(* IEC 61131-3 sources: CS_4_Aufzugsteuerung/src/Stations/CP112/Steuerung/Class/_DriveAxisBase (part 2) *)

      16#1B: //27-> PWM setvalue for G-MODE=7 + controlword
        //PWM from -1000 to 1000 for -100% to 100% is preset via SetSpeed
        SyncPara.SetSpeed.size := 2;
        SyncPara.SetSpeed.ptr := #SetValuePtr^.a_SyncValues[x];
        SyncPara.SetSpeed.userinfo := 1;

        SyncPara.ControlWord.size := 2;
        SyncPara.ControlWord.ptr := #SetValuePtr^.a_SyncValues[x] + sizeof(UINT);
        SyncPara.ControlWord.userinfo := 0;

        SyncPara.SetTorque.size := 2;
        SyncPara.SetTorque.ptr := #SetValuePtr^.a_SyncValues[x] + sizeof(UINT);
        SyncPara.SetTorque.userinfo := 0;

    end_case;

  end_for;

END_FUNCTION

FUNCTION VIRTUAL GLOBAL _DriveAxisBase::SetPos::Write
	VAR_INPUT
		input (EAX) 	: DINT;
	END_VAR
	VAR_OUTPUT
		result (EAX) 	: DINT;
	END_VAR

  if (SyncPara.SetPos.ptr <> NIL) & bOnlineFinished then
    SetPos:=input;
    SyncPara.SetPos.ptr^:=input;
  end_if;

 	result := SetPos;

END_FUNCTION

FUNCTION VIRTUAL GLOBAL _DriveAxisBase::SetSpeed::Write
	VAR_INPUT
		input (EAX) 	: DINT;
	END_VAR
	VAR_OUTPUT
		result (EAX) 	: DINT;
	END_VAR

	if bOnlineFinished then
    SetSpeed := Write_SetSpeed(input);  //write value to PDO data, and set possible statusflags.
        end_if;
 	result := SetSpeed;

END_FUNCTION

FUNCTION VIRTUAL GLOBAL _DriveAxisBase::SetCurrent::Write
	VAR_INPUT
		input (EAX) 	: DINT;
	END_VAR
	VAR_OUTPUT
		result (EAX) 	: DINT;
	END_VAR

  if (SyncPara.SetCurrent.ptr <> NIL) & bOnlineFinished then
    SetCurrent:=input;
    if (SyncPara.SetCurrent.size=4) then
      SyncPara.SetCurrent.ptr^:=input;
    elsif (SyncPara.SetCurrent.size=2) then
      if SyncPara.SetCurrent.userinfo = 1 then
        SyncPara.SetCurrent.ptr^$INT:=to_int(input / 10); //because we always get mA and in one case we must send cA
      else
        SyncPara.SetCurrent.ptr^$INT:=to_int(input); //32-Bit-Steuerwort
      end_if;
    end_if;
  end_if;

  result := SetCurrent;

END_FUNCTION

FUNCTION VIRTUAL GLOBAL _DriveAxisBase::ControlWord::Write
	VAR_INPUT
		input (EAX) 	: DS402_Control;
	END_VAR
	VAR_OUTPUT
		result (EAX) 	: DS402_Control;
	END_VAR
  VAR
  	cBuffer : BDINT; //ControlWord Buffer
  END_VAR

  cBuffer := 0; // local variable

  if (SyncPara.ControlWord.ptr <> NIL) & bOnlineFinished then

    if (SyncPara.ControlWord.userinfo=0) then //normal controlword

      cBuffer.1  :=input.EnableOperation;   //DRIVE ENABLE
      cBuffer.2  :=input.ResetFault;        //FAULT RESET
      cBuffer.3  :=input.ManufactureSpec1;  //AMODE2
      cBuffer.4  :=input.ManufactureSpec2;  //KFBRW3
      cBuffer.5  :=input.ManufactureSpec4;  //Output1
      cBuffer.6  :=input.ManufactureSpec5;  //Output2
      cBuffer.7  :=input.ManufactureSpec3;  //KBRAKE
      cBuffer.8  :=input.Reserved1;         //ECHO
      cBuffer.9  :=input.OperationModeSpec1;//SINGLE CAPTURE

      cBuffer:=TorqueCalculation(cBuffer, AxTorqueControl); //cBuffer -> we must add TorqueControl

      SyncPara.ControlWord.ptr^$INT:=to_int(cBuffer);

    elsif(SyncPara.ControlWord.userinfo=1)then

      cBuffer.1 :=input.SwitchOn;
      cBuffer.2 :=input.EnableVoltage;
      cBuffer.3 :=input.QuickStop;
      cBuffer.4 :=input.EnableOperation;    //DRIVE ENABLE
      cBuffer.5 :=input.OperationModeSpec1;
      cBuffer.6 :=input.OperationModeSpec2;
      cBuffer.7 :=input.OperationModeSpec3;
      cBuffer.8 :=input.ResetFault;         //FAULT RESET
      cBuffer.9 :=input.Halt;
      cBuffer.10 :=input.Reserved1;
      cBuffer.11 :=input.Reserved2;
      cBuffer.12 :=input.ManufactureSpec1;  //AMODE2
      cBuffer.13 :=input.ManufactureSpec2;  //KFBRW3
      cBuffer.14 :=input.ManufactureSpec3;  //KBRAKE
      cBuffer.15 :=input.ManufactureSpec4;  //Output1
      cBuffer.16 :=input.ManufactureSpec5;  //Output2

      SyncPara.ControlWord.ptr^$INT:=to_int(cBuffer);

    end_if;

  end_if;

  ControlWord := input;
  result := ControlWord;

END_FUNCTION

FUNCTION VIRTUAL GLOBAL _DriveAxisBase::AxEnable::Write
	VAR_INPUT
		input (EAX) 	: DINT;
	END_VAR
	VAR_OUTPUT
		result (EAX) 	: DINT;
	END_VAR

  if (SyncPara.ControlWord.ptr <> NIL) & bOnlineFinished then
    AxEnable:= Write_Enable( input AND 1 );
  end_if;
  result:=AxEnable;

END_FUNCTION

FUNCTION VIRTUAL GLOBAL _DriveAxisBase::AxErrorQuit::Write
	VAR_INPUT
		input (EAX) 	: DINT;
	END_VAR
	VAR_OUTPUT
		result (EAX) 	: DINT;
	END_VAR

  if SyncPara.ControlWord.ptr & (FirstErrorReset = 0) & bOnlineFinished then

    if (AxError = 1) then

      ErrorQuitHandling(input);

    end_if;

  end_if;

  result := AxErrorQuit;

END_FUNCTION

FUNCTION VIRTUAL GLOBAL _DriveAxisBase::AxTorqueControl::Write
	VAR_INPUT
		input (EAX) 	: UDINT;
	END_VAR
	VAR_OUTPUT
		result (EAX) 	: UDINT;
	END_VAR

  if (SyncPara.SetTorque.ptr <> NIL) & bOnlineFinished then
    SetAxTorque(input);
  end_if;

  result := AxTorqueControl;

END_FUNCTION

FUNCTION _DriveAxisBase::TorqueCalculation
	VAR_INPUT
		cBuffer 	: BDINT;
		input 	  : UDINT;
	END_VAR
	VAR_OUTPUT
		result 	  : BDINT;
	END_VAR
  VAR
  	IReduce   : UDINT;
  END_VAR

  IReduce := ((DRIVEAXIS_TORQUE_LIMITATION_VALUE - input) * 63) / DRIVEAXIS_TORQUE_LIMITATION_VALUE; // calculate the bits for the current reducing

  IReduce := IReduce SHL 10 ;
  cBuffer := cBuffer AND 16#3FF;
  cBuffer+=IReduce$BDINT;

  result:=cBuffer;

END_FUNCTION

//****************************************************************************************************\\
//**################################################################################################**\\
//**************************** everything for getting the actual values!! ****************************\\
//**################################################################################################**\\
//****************************************************************************************************\\

FUNCTION VIRTUAL GLOBAL _DriveAxisBase::GetSynchronPara
  VAR
  	x:SINT;
    SetAVALTT:HSINT;
  END_VAR

  ActValuePtr := DriveMng.GetAxisRdPtr(usAxisIndex); // Zeiger auf die Sollwerte von der Struktur t_ReadValuePtr

  for x:=4 to 0 by -1 do
    SetAVALTT:=ActValues[x];

    case SetAVALTT of

      16#01: //1 -> I-N
        SyncPara.ActSpeed.ptr:=#ActValuePtr^.a_SyncValues[x];
        SyncPara.ActSpeed.size:=4;
        SyncPara.ActSpeed.userinfo:=0;

      16#02: //2 -> I-NFILT
        SyncPara.ActSpeed.ptr:=#ActValuePtr^.a_SyncValues[x];
        SyncPara.ActSpeed.size:=4;
        SyncPara.ActSpeed.userinfo:=0;

//      16#03:
//
//        SyncPara.SetPos

      16#05: //5 -> I-IQ
        SyncPara.ActCurrent.ptr:=#ActValuePtr^.a_SyncValues[x];
        SyncPara.ActCurrent.size:=4;
        SyncPara.ActCurrent.userinfo:=0;

      16#07: //7 -> I-POS
        SyncPara.ActPos.ptr:=#ActValuePtr^.a_SyncValues[x];
        SyncPara.ActPos.size:=4;
        SyncPara.ActPos.userinfo:=0;

      16#09: //9 -> I-PE
        SyncPara.Xw.ptr:=#ActValuePtr^.a_SyncValues[x];
        SyncPara.Xw.size:=4;
        SyncPara.Xw.userinfo:=0;

      16#0A: //10 -> I-IQ + stateword (cA!)
        SyncPara.ActCurrent.ptr:=#ActValuePtr^.a_SyncValues[x];
        SyncPara.ActCurrent.size:=2;
        SyncPara.ActCurrent.userinfo:=1;

        SyncPara.StateWord.ptr:=#ActValuePtr^.a_SyncValues[x]+sizeof(UINT);
        SyncPara.StateWord.size:=2;
        SyncPara.StateWord.userinfo:=0;

      16#0E: //14 -> I-PE + stateword
        SyncPara.Xw.ptr:=#ActValuePtr^.a_SyncValues[x];
        SyncPara.Xw.size:=2;
        SyncPara.Xw.userinfo:=0;

        SyncPara.StateWord.ptr:=#ActValuePtr^.a_SyncValues[x]+sizeof(UINT);
        SyncPara.StateWord.size:=2;
        SyncPara.StateWord.userinfo:=0;

      16#14: //20 -> Current in Promille + stateword
        SyncPara.ActCurrent.ptr:=#ActValuePtr^.a_SyncValues[x];
        SyncPara.ActCurrent.size:=2;
        SyncPara.ActCurrent.userinfo:=0;

        SyncPara.StateWord.ptr:=#ActValuePtr^.a_SyncValues[x]+sizeof(UINT);
        SyncPara.StateWord.size:=2;
        SyncPara.StateWord.userinfo:=1;

      16#15: //21 -> I-POS 2 position of optional encoder
        if (SyncPara.ActPos.ptr = NIL) then
          SyncPara.ActPos.ptr:=#ActValuePtr^.a_SyncValues[x];
          SyncPara.ActPos.size:=4;
          SyncPara.ActPos.userinfo:=0;
        end_if;

      16#17: //23 -> digital inputs + stateword
        SyncPara.DigInputs.ptr:=#ActValuePtr^.a_SyncValues[x];
        SyncPara.DigInputs.size:=8; //no inputs
        SyncPara.DigInputs.userinfo:=0;

        SyncPara.StateWord.ptr:=#ActValuePtr^.a_SyncValues[x]+sizeof(UINT);
        SyncPara.StateWord.size:=2;
        SyncPara.StateWord.userinfo:=0;

      16#1C: //28 -> MultiTurn Pos VSDC151
        SyncPara.ActPos.ptr:=#ActValuePtr^.a_SyncValues[x];
        SyncPara.ActPos.size:=4;
        SyncPara.ActPos.userinfo:=0;

    end_case;

  end_for;

END_FUNCTION

FUNCTION VIRTUAL GLOBAL _DriveAxisBase::ActPos::Read
	VAR_OUTPUT
		output (EAX) 	: DINT;
	END_VAR

  if (SyncPara.ActPos.ptr <> NIL) & bOnlineFinished then
    ActPos:=SyncPara.ActPos.ptr^;
  else
    ActPos:=0;
  end_if;

  output := ActPos;

END_FUNCTION

FUNCTION VIRTUAL GLOBAL _DriveAxisBase::ActSpeed::Read
	VAR_OUTPUT
		output (EAX) 	: DINT;
	END_VAR

  if (SyncPara.ActSpeed.ptr <> NIL) & bOnlineFinished then
    ActSpeed:=SyncPara.ActSpeed.ptr^;
  else
    ActSpeed:=0;
  end_if;

  output := ActSpeed;

END_FUNCTION

FUNCTION VIRTUAL GLOBAL _DriveAxisBase::ActCurrent::Read
	VAR_OUTPUT
		output (EAX) 	: DINT;
	END_VAR

  if (SyncPara.ActCurrent.ptr <> NIL) & bOnlineFinished then
    if SyncPara.ActCurrent.size = 4 then
      ActCurrent:=SyncPara.ActCurrent.ptr^;

    elsif SyncPara.ActCurrent.size = 2 then
      if SyncPara.ActCurrent.userinfo = 1 then
        ActCurrent := to_dint(SyncPara.ActCurrent.ptr^$INT) * 10; //because we want to see mA and not cA
      else
        ActCurrent := to_dint(SyncPara.ActCurrent.ptr^$INT);
      end_if;
    end_if;
  else
    ActCurrent:=0;
  end_if;

  output := ActCurrent;

END_FUNCTION

FUNCTION VIRTUAL GLOBAL _DriveAxisBase::ActXw::Read
	VAR_OUTPUT
		output (EAX) 	: DINT;
	END_VAR

  if (SyncPara.Xw.ptr <> NIL) & bOnlineFinished then
    if SyncPara.Xw.size = 4 then
      ActXw:=SyncPara.Xw.ptr^;
    elsif SyncPara.Xw.size = 2 then
      ActXw := to_dint(SyncPara.Xw.ptr^$INT);
    end_if;
  else
    ActXw:=0;
  end_if;

  output := ActXw;

END_FUNCTION

FUNCTION VIRTUAL GLOBAL _DriveAxisBase::StateWord::Read
	VAR_OUTPUT
		output (EAX) 	: DS402_State;
	END_VAR
  VAR
  	sBuffer : BDINT; //StateWord Buffer
  END_VAR

  if (SyncPara.StateWord.ptr <> NIL) & bOnlineFinished then
    sBuffer := SyncPara.StateWord.ptr^$BDINT; //normales Statuswort

    if (SyncPara.StateWord.userinfo=0) then
      StateWord.ReadyToSwitchOn     :=  sBuffer.1;  //READY TO SWITCH ON
      StateWord.SwitchedOn          :=  sBuffer.2;  //EXT ENABLE LOCKED&ENABLE
      StateWord.OperationEnabled    :=  sBuffer.3;  //OPERATION_ENABLE
      StateWord.Fault               :=  sBuffer.4;  //ERROR
      StateWord.Warning             :=  sBuffer.5;  //WARNING
      StateWord.Remote              :=  sBuffer.6;  //PLL Bit0
      StateWord.VoltageEnabled      :=  sBuffer.7;  //PLL Bit1
      StateWord.SwitchOnDisabled    :=  sBuffer.8;  //ECHO
      StateWord.OperationModeSpec1  :=  sBuffer.9;  //Capture Toggle Bit (I-CAP)
      StateWord.OperationModeSpec2  :=  sBuffer.10; //Capture 4 Toggle Bit (I-CAP4)
      StateWord.InternalLimitActive :=  sBuffer.11; //MULTITURN REVOLUTION ERROR
      StateWord.ManufactureSpec1    :=  sBuffer.12; //Digital Input 1
      StateWord.ManufactureSpec2    :=  sBuffer.13; //Digital Input 2
      StateWord.ManufactureSpec3    :=  sBuffer.14; //Digital Input 3
      StateWord.QuickStop           :=  sBuffer.15; //Digital Input 4
      StateWord.TargetReached       :=  sBuffer.16; //Digital Input 5

    elsif(SyncPara.StateWord.userinfo=1) then
      StateWord.ReadyToSwitchOn     :=  sBuffer.1;  //READY TO SWITCH ON
      StateWord.SwitchedOn          :=  sBuffer.2;  //EXT.ENABLE=LOCKED&ENABLE
      StateWord.OperationEnabled    :=  sBuffer.3;  //OPERATION_ENABLE
      StateWord.Fault               :=  sBuffer.4;  //ERROR
      StateWord.Warning             :=  sBuffer.5;  //WARNING
      StateWord.QuickStop           :=  sBuffer.6;
      StateWord.SwitchOnDisabled    :=  sBuffer.7;
      StateWord.VoltageEnabled      :=  sBuffer.8;
      StateWord.ManufactureSpec1    :=  sBuffer.9;
      StateWord.ManufactureSpec2    :=  sBuffer.10;
      StateWord.TargetReached       :=  sBuffer.11;
      StateWord.ManufactureSpec3    :=  sBuffer.12;
      StateWord.OperationModeSpec1  :=  sBuffer.13;
      StateWord.OperationModeSpec2  :=  sBuffer.14;
      StateWord.Remote              :=  sBuffer.15; //PLL nicht eingerastet
      StateWord.InternalLimitActive :=  sBuffer.16; //MULTITURN REVOLUTION ERROR
    end_if;

  else
    StateWord := 0;
  end_if;

  output := StateWord;

END_FUNCTION

FUNCTION VIRTUAL GLOBAL _DriveAxisBase::AxError::Read
	VAR_OUTPUT
		output (EAX) : DINT;
	END_VAR

  //Error of Axis gets only shown, if Axis is Online
  if bOnlineFinished then
    AxError := GetAxError();
  else
    AxError := 0;
  end_if;

  output := AxError;

END_FUNCTION

FUNCTION _DriveAxisBase::LoadDrivePara
  VAR
    pTabAdress : ^DINT;
    TabLength   : DINT;
  END_VAR

  // load the parameter data to the para objects
  case DriveInitType of

    _SDDSTDTABLE :

     pTabAdress := GetTabAdress(TabType:= 0, bdSettings.bSendMPara, #TabLength);
     SetListToParObj(pData:= (pTabAdress)$^DINT, udLen:=TabLength$UDINT);

    _SDDL2TABLE :
    // load the data of the table
      pTabAdress := GetTabAdress(TabType:= 1, bdSettings.bSendMPara, #TabLength);
      SetListToParObj(pData:= (pTabAdress)$^DINT, udLen:=TabLength$UDINT);

    _SDDRAMEX,
    _SDDFILE :
      pSDDData$^void := DriveAxisSet.GetMemPtr();
      if pSDDData <> NIL then
        // load the data of the memory
        SetListToParObj(pData:= (pSDDData$DINT + pSDDData^.AxOffset)$^DINT, udLen:=pSDDData^.AxLength);
      end_if;

  end_case;

END_FUNCTION

FUNCTION _DriveAxisBase::SetListToParObj
	VAR_INPUT
		pData 	: ^DINT;
		udLen 	: UDINT;
	END_VAR
	VAR_OUTPUT
		retcode 	: BOOL;
	END_VAR
  VAR
    pHlp          : ^DINT;
    x             : UDINT;
    pThisNewInst  : ^void;
    usParaNr      : USINT;
    ParaValue     : DINT;
    UserPara      : CmdStruct;
    UserResult    : Results;
  END_VAR

  retcode := FALSE;

  //hier konnte es zu einem Problem kommen kann wenn pThisNewInst nicht init war.
  pThisNewInst := NIL; //BleErn 19.08.2010 11:27

  if (bdSettings.bAxSetPara = FALSE) | (pData = NIL) then
    return;
  end_if;

  x := 0;
  pHlp := pData;

  while x < udLen do

    usParaNr := pHlp^$USINT;
    pHlp += sizeof(USINT);
    x += sizeof(USINT);

    if usParaNr <= MAX_MOTOR_PARA then
      pThisNewInst$DINT := AxSetPara[IDX_MOTOR_PARA];
    elsif usParaNr <= MAX_DRIVE_PARA then
      pThisNewInst$DINT := AxSetPara[IDX_DRIVE_PARA];
    elsif usParaNr <= MAX_CURRENT_PARA then
      pThisNewInst$DINT := AxSetPara[IDX_CURRENT_PARA];
    elsif usParaNr <= MAX_VEL_PARA then
      pThisNewInst$DINT := AxSetPara[IDX_VEL_PARA];
    elsif usParaNr <= MAX_POS_PARA then
      pThisNewInst$DINT := AxSetPara[IDX_POS_PARA];
    elsif usParaNr <= MAX_FD_PARA then
      pThisNewInst$DINT := AxSetPara[IDX_FD_PARA];
    elsif usParaNr <= MAX_APPLI_PARA then
      pThisNewInst$DINT := AxSetPara[IDX_APPLI_PARA];
    elsif usParaNr <= MAX_ERRORHANDLING then
      pThisNewInst$DINT := AxSetPara[IDX_ERRORHANDLING];
    end_if;

    ParaValue := pHlp^$DINT;
    if pThisNewInst <> NIL then
      UserPara.uiCmd := SDD_REFRESH_SETPARA;
      UserPara.aPara[0] := to_dint(usParaNr);
      UserPara.aPara[1] := ParaValue;
      pThisNewInst$^VirtualBase^.NewInst(#UserPara, #UserResult);
    end_if;

    pHlp += sizeof(UDINT);
    x += sizeof(UDINT);

  end_while;

END_FUNCTION

FUNCTION VIRTUAL GLOBAL _DriveAxisBase::SDDProcess
  VAR
    tmpStr : array [0..20] of char;
    retcode : iprStates;
    dError : DINT;
  END_VAR

  //SA 23391 - ObeChr: Wait for Online before starting SDDCmdInterface
  if Online = 1 then

    case SDDCmdIntfc of

    _SDDIDLE :
      // do nothing

    _SDDREADALL :
      if bdSettings.bStartRead = FALSE then
        bdSettings.bStartRead := TRUE;
        // check if a read is possible
        if ChkParaRead(0) = FALSE then
          SDDCmdIntfc := _SDDIDLE;
        else
          ParaReadProc();
        end_if;
      else
        // überprüfen ob alle Parameter schon vorhanden sind
        ParaReadProc();
        if (bdSettings.bReadAxFin = TRUE) then
          SDDCmdIntfc := _SDDIDLE;
          bdSettings.bStartRead := FALSE;
        end_if;
      end_if;

    _SDDINIT :

      if (AxEnable = 0)  then
        if OldSDDCmdIntfc <> SDDCmdIntfc then
          DriveMng.InitDrive(0); // start the initialisation of the drive
          Init_Again:=true;
          //bdSettings.bDriveInitialized:=true;
        end_if;
      else
        SDDCmdIntfc := _SDDIDLE;
      end_if;

    _SDDURINIT :

      if (AxEnable = 0) then
        if OldSDDCmdIntfc <> SDDCmdIntfc then
          DriveMng.InitDrive(1); // start the initialisation of the drive
          InitASyncPara(); // initialize the structure
          Init_Again:=true;
        end_if;
      else
        SDDCmdIntfc := _SDDIDLE;
      end_if;

    _SDDEXDATA,
    _SDDEXDATAXML:

      // only if a object of the correct class is connected
      if DriveAxisSet.ChkFileHandle() then

        if OldSDDCmdIntfc <> SDDCmdIntfc then
          pSDDData$^void := DriveAxisSet.GetMemPtr();

          // Always Call SetDriveType incause GetDriveTypeStr fails or an older Version of _DriveFileHandling is used
          DriveAxisSet.SetDriveType(eDriveType:=GetDriveType());

          _strcpy(#pSDDData^.AxName[0],#szObjName[0]); //here the name of the object is set to the struct

          // Set tmpStr to 0 incase GetDriveTypeStr does not return a valid string.
          tmpStr[0] := 0;
          DriveMng.GetDriveTypeStr(eDriveType:=GetDriveType(), pDriveTypeStr:=#tmpStr[0], DriveTypeStrSize:=sizeof(tmpStr) );
          if tmpStr[0] then
            DriveAxisSet.SetDriveTypeStr(pDriveTypeStr:= #tmpStr[0]);
          end_if;
          DriveAxisSet.SetUserSSDCmd(SDDCmdIntfc, pSDDData);

        else
          SDDCmdIntfc := DriveAxisSet.GetUserSSDCmd();
        end_if;
      else
        LogError(pMsg:="@06F3 (_DriveAxisBase::SDDProcess) Failed export drive parameters. Check if client 'FileHandle' is connected.");
        SDDCmdIntfc := _SDDERROR;
      end_if;

    _SDDIMDATAXML:

      if DriveAxisSet.ChkFileHandle() then

        if OldSDDCmdIntfc <> SDDCmdIntfc then
          pSDDData$^void := DriveAxisSet.GetMemPtr();

          _strcpy(#pSDDData^.AxName[0],#szObjName[0]); //here the name of the object is set to the struct
          DriveAxisSet.SetUserSSDCmd(SDDCmdIntfc, pSDDData);

        else

          if DriveAxisSet.GetUserSSDCmd() = _SDDIDLE then
            // Read xml file done

            // Insert Crc into the imported Data
            pSDDData^.udCRC32 := DriveAxisSet.CalcCRC32((pSDDData + sizeof(UDINT))$^UDINT, pSDDData^.udLen - sizeof(UDINT));

            // now save all parameters in the SRAM / FILE
            if DriveInitType = _SDDRAMEX then
              pSDDData$^void := DriveAxisSet.GetMemPtr();
              DriveAxisSet.SaveRamExData(pData:= pSDDData, udLen:= pSDDData^.udLen, udOffset:= 0);

            elsif DriveInitType = _SDDFILE then
              pSDDData$^void := DriveAxisSet.GetMemPtr();
              DriveAxisSet.SaveRamFileData(pData:= pSDDData, udLen:= pSDDData^.udLen, udOffset:= 0);

            end_if;

            // Use _SDDINIT to tranfer Parametera from ramfile/sram to drive
            SDDCmdIntfc := _SDDINIT;  // Set after SaveRamExData, SaveRamFileData because Filehandling may suspend task

            return; // Return needed here so that _SDDINIT is registered as a new command
          end_if;

        end_if;
      else
        LogError(pMsg:="@06F5 (_DriveAxisBase::SDDProcess) Failed import drive parameters. Check if client 'FileHandle' is connected.");
        SDDCmdIntfc := _SDDERROR;
      end_if;

      _SDDEXLOGFILE:

        // First call since SDDCmdIntfc was set.
        if OldSDDCmdIntfc <> SDDCmdIntfc then

          retcode := DriveMng.GetLogFile(pDestinationDPNE:=NIL, pdError:=#dError);

          if retcode = ERROR then

            LogValue("@0846 (_DriveAxisBase::SDDProcess) Failed to start read logfile. Error code: -0x{0}", (-dError)$UDINT);
            SDDCmdIntfc := _SDDERROR;

          end_if;

        else

          retcode := DriveMng.GetFileState(pdError:=#dError);

          if retcode = READY then

            SDDCmdIntfc := _SDDIDLE;

          elsif retcode = ERROR then

            LogValue("@0847 (_DriveAxisBase::SDDProcess) Failed read logfile. Error code: -0x{0}", (-dError)$UDINT);
            SDDCmdIntfc := _SDDERROR;

          end_if;

        end_if;

    end_case;

    OldSDDCmdIntfc := SDDCmdIntfc;

  end_if;

END_FUNCTION

FUNCTION VIRTUAL GLOBAL _DriveAxisBase::SDDCmdIntfc::Write
	VAR_INPUT
		input (EAX) 	: _SDDUSERCMD;
	END_VAR
	VAR_OUTPUT
		result (EAX) 	: _SDDUSERCMD;
	END_VAR

  if ((SDDCmdIntfc = _SDDIDLE) |
      (SDDCmdIntfc = _SDDERROR)) then
    SDDCmdIntfc := input;
    result := SDDCmdIntfc;
  else
    result$DINT := ACCESS_DENIED;
  end_if;

END_FUNCTION

FUNCTION _DriveAxisBase::ChkParaRead
	VAR_INPUT
		ChkType 	: DINT;
	END_VAR
	VAR_OUTPUT
		retcode 	: BOOL;
	END_VAR

  retcode := FALSE;

  case ChkType of
  0 : // check if a reading command is allowed

    bdSettings.bReadAx := FALSE;

    bdSettings.bReadAxFin := FALSE;

    if (bdSettings.bAxSetPara = TRUE)then
      bdSettings.bReadAx := TRUE;
      ParaReadCmdAx := 1;
      retcode := TRUE;
    else
      bdSettings.bReadAxFin := TRUE;
    end_if;

  1 : // check if we can send the next reading commands
    if ParaReadCmdAx = 2 then
      if AxASyncPara.ActEntries < 10 then
        retcode := TRUE;
      end_if;
    end_if;

  end_case;

END_FUNCTION

FUNCTION _DriveAxisBase::ParaReadProc
  VAR
    dValue      : DINT;
    pThis       : ^void;
    i           : DINT;
    UserPara    : CmdStruct;
    UserResult  : Results;
  END_VAR
        // Start laden aller Parameter vom Drive
        // folgender Ablauf :
        // 1. Es wird für jede Achse die Anforderung in den Ringbuffer geschrieben (30mal).(Eigene Kennung erforderlich ?);
        // 2. Warten bis nur mehr 10 Einträge vorhanden sind, und dann die nächsten Einträge absetzen
        // 3. wenn alle Einträge abgesetzt sind, (letzter Eintrag muss eine extra Kennung haben), wird überprüft wann alle Daten vorhanden sind
        // 4. Wenn ein Wert eines Parameters ankommt, wird dieser in den Speicher geschrieben, dies ist abhängig von der Sicherungsauswahl. Ist eine Tabelle ausgewählt
        //    werden die Daten sofort an die Parameterklassen gesendet, sind keine Parameterobjekte vorhanden, so wird der Vorgang gar nicht durchgeführt.
        // 5. Wenn der letzte Wert des Parameters kommt, wird die Chksumme neu berechnet, die Daten weggesichert, und die Parameterobjekte aktualisiert

  dValue := 0;

 if bdSettings.bReadAx = TRUE then
    case ParaReadCmdAx of

    0 : //idle step

    1 : // set the first entries in the buffer
      // set the info busy to all para classes
      UserPara.uiCmd := SDD_ASYNC_BUSY;

      for i := IDX_MOTOR_PARA to IDX_ERRORHANDLING do
        pThis$DINT := AxSetPara[i];
        if pThis <> NIL then
          // Set the state BUSY
          pThis$^VirtualBase^.NewInst(#UserPara, #UserResult);
        end_if;
      end_for;

      if AxSetPara[IDX_MOTOR_PARA] <> 0 then
        pThis$DINT := AxSetPara[IDX_MOTOR_PARA];

        AddASyncEntry(usParaNr:= SDD_M_NAME1, usRdWr:= 0, dValue:= dValue, pThisObj:= pThis, usEntry:= 1);
        AddASyncEntry(usParaNr:= SDD_M_NAME2, usRdWr:= 0, dValue:= dValue, pThisObj:= pThis, usEntry:= 1);
        AddASyncEntry(usParaNr:= SDD_M_NAME3, usRdWr:= 0, dValue:= dValue, pThisObj:= pThis, usEntry:= 1);
        AddASyncEntry(usParaNr:= SDD_M_INULL, usRdWr:= 0, dValue:= dValue, pThisObj:= pThis, usEntry:= 1);
        AddASyncEntry(usParaNr:= SDD_M_IPEAK, usRdWr:= 0, dValue:= dValue, pThisObj:= pThis, usEntry:= 1);
        AddASyncEntry(usParaNr:= SDD_M_NMAX, usRdWr:= 0, dValue:= dValue, pThisObj:= pThis, usEntry:= 1);
        AddASyncEntry(usParaNr:= SDD_M_POL, usRdWr:= 0, dValue:= dValue, pThisObj:= pThis, usEntry:= 1);
        AddASyncEntry(usParaNr:= SDD_M_TORQUE, usRdWr:= 0, dValue:= dValue, pThisObj:= pThis, usEntry:= 1);
        AddASyncEntry(usParaNr:= SDD_M_L, usRdWr:= 0, dValue:= dValue, pThisObj:= pThis, usEntry:= 1);
        AddASyncEntry(usParaNr:= SDD_M_R, usRdWr:= 0, dValue:= dValue, pThisObj:= pThis, usEntry:= 1);
        AddASyncEntry(usParaNr:= SDD_M_J, usRdWr:= 0, dValue:= dValue, pThisObj:= pThis, usEntry:= 1);
        AddASyncEntry(usParaNr:= SDD_M_TYPE, usRdWr:= 0, dValue:= dValue, pThisObj:= pThis, usEntry:= 1);
        AddASyncEntry(usParaNr:= SDD_M_RPOL, usRdWr:= 0, dValue:= dValue, pThisObj:= pThis, usEntry:= 1);
        AddASyncEntry(usParaNr:= SDD_M_ROFF, usRdWr:= 0, dValue:= dValue, pThisObj:= pThis, usEntry:= 1);
        AddASyncEntry(usParaNr:= SDD_M_RPULSE, usRdWr:= 0, dValue:= dValue, pThisObj:= pThis, usEntry:= 1);
        AddASyncEntry(usParaNr:= SDD_M_RTEMP, usRdWr:= 0, dValue:= dValue, pThisObj:= pThis, usEntry:= 1);
        AddASyncEntry(usParaNr:= SDD_M_SER, usRdWr:= 0, dValue:= dValue, pThisObj:= pThis, usEntry:= 1);
        AddASyncEntry(usParaNr:= SDD_M_BRAKE, usRdWr:= 0, dValue:= dValue, pThisObj:= pThis, usEntry:= 1);
        AddASyncEntry(usParaNr:= SDD_M_IFWEAK, usRdWr:= 0, dValue:= dValue, pThisObj:= pThis, usEntry:= 1);
        AddASyncEntry(usParaNr:= SDD_M_BRDIS, usRdWr:= 0, dValue:= dValue, pThisObj:= pThis, usEntry:= 1);
        AddASyncEntry(usParaNr:= SDD_M_BREN, usRdWr:= 0, dValue:= dValue, pThisObj:= pThis, usEntry:= 1);
        AddASyncEntry(usParaNr:= SDD_M_IMAG, usRdWr:= 0, dValue:= dValue, pThisObj:= pThis, usEntry:= 1);
        AddASyncEntry(usParaNr:= SDD_M_TROT, usRdWr:= 0, dValue:= dValue, pThisObj:= pThis, usEntry:= 1);
        AddASyncEntry(usParaNr:= SDD_M_UN, usRdWr:= 0, dValue:= dValue, pThisObj:= pThis, usEntry:= 1);
        AddASyncEntry(usParaNr:= SDD_M_UBOOST, usRdWr:= 0, dValue:= dValue, pThisObj:= pThis, usEntry:= 1);
        AddASyncEntry(usParaNr:= SDD_M_KN, usRdWr:= 0, dValue:= dValue, pThisObj:= pThis, usEntry:= 1);
      end_if;

      if AxSetPara[IDX_DRIVE_PARA] <> 0 then
        pThis$DINT := AxSetPara[IDX_DRIVE_PARA];
        AddASyncEntry(usParaNr:= SDD_G_MODE, usRdWr:= 0, dValue:= dValue, pThisObj:= pThis, usEntry:= 1);
        AddASyncEntry(usParaNr:= SDD_G_CETIME, usRdWr:= 0, dValue:= dValue, pThisObj:= pThis, usEntry:= 1);
        AddASyncEntry(usParaNr:= SDD_G_VMAINS, usRdWr:= 0, dValue:= dValue, pThisObj:= pThis, usEntry:= 1);
        AddASyncEntry(usParaNr:= SDD_G_VBUSM, usRdWr:= 0, dValue:= dValue, pThisObj:= pThis, usEntry:= 1);
        AddASyncEntry(usParaNr:= SDD_G_VBUSM, usRdWr:= 0, dValue:= dValue, pThisObj:= pThis, usEntry:= 1);
        AddASyncEntry(usParaNr:= SDD_G_MTEMPK, usRdWr:= 0, dValue:= dValue, pThisObj:= pThis, usEntry:= 1);
        AddASyncEntry(usParaNr:= SDD_G_MTEMPE, usRdWr:= 0, dValue:= dValue, pThisObj:= pThis, usEntry:= 1);
        AddASyncEntry(usParaNr:= SDD_G_PWM, usRdWr:= 0, dValue:= dValue, pThisObj:= pThis, usEntry:= 1);
        AddASyncEntry(usParaNr:= SDD_G_DELAY, usRdWr:= 0, dValue:= dValue, pThisObj:= pThis, usEntry:= 1);
        AddASyncEntry(usParaNr:= SDD_G_FTEMP, usRdWr:= 0, dValue:= dValue, pThisObj:= pThis, usEntry:= 1);
        AddASyncEntry(usParaNr:= SDD_G_EMRAMP, usRdWr:= 0, dValue:= dValue, pThisObj:= pThis, usEntry:= 1);
        AddASyncEntry(usParaNr:= SDD_G_MASKE1, usRdWr:= 0, dValue:= dValue, pThisObj:= pThis, usEntry:= 1);
        AddASyncEntry(usParaNr:= SDD_G_MASKE2, usRdWr:= 0, dValue:= dValue, pThisObj:= pThis, usEntry:= 1);
        AddASyncEntry(usParaNr:= SDD_G_MASKW, usRdWr:= 0, dValue:= dValue, pThisObj:= pThis, usEntry:= 1);
        AddASyncEntry(usParaNr:= SDD_G_MASKD, usRdWr:= 0, dValue:= dValue, pThisObj:= pThis, usEntry:= 1);
        AddASyncEntry(usParaNr:= SDD_G_VRAMP, usRdWr:= 0, dValue:= dValue, pThisObj:= pThis, usEntry:= 1);
        AddASyncEntry(usParaNr:= SDD_G_SRAMP, usRdWr:= 0, dValue:= dValue, pThisObj:= pThis, usEntry:= 1);
        AddASyncEntry(usParaNr:= SDD_G_RBAL, usRdWr:= 0, dValue:= dValue, pThisObj:= pThis, usEntry:= 1);
      end_if;

      ParaReadCmdAx := 2;

    2 :
      // wait until only 10 entries in the buffer

      if ChkParaRead(ChkType:= 1) = TRUE then
        ParaReadCmdAx := 3;
      end_if;

    3 :
      // send the rest

      if AxSetPara[IDX_CURRENT_PARA] <> 0 then
        pThis$DINT := AxSetPara[IDX_CURRENT_PARA];
        AddASyncEntry(usParaNr:= SDD_C_KPQ, usRdWr:= 0, dValue:= dValue, pThisObj:= pThis, usEntry:= 1);
        AddASyncEntry(usParaNr:= SDD_C_TN, usRdWr:= 0, dValue:= dValue, pThisObj:= pThis, usEntry:= 1);
        AddASyncEntry(usParaNr:= SDD_C_KDREL, usRdWr:= 0, dValue:= dValue, pThisObj:= pThis, usEntry:= 1);
        AddASyncEntry(usParaNr:= SDD_C_KPDREL, usRdWr:= 0, dValue:= dValue, pThisObj:= pThis, usEntry:= 1);
        AddASyncEntry(usParaNr:= SDD_C_KPNULL, usRdWr:= 0, dValue:= dValue, pThisObj:= pThis, usEntry:= 1);
        AddASyncEntry(usParaNr:= SDD_C_KPPEAK, usRdWr:= 0, dValue:= dValue, pThisObj:= pThis, usEntry:= 1);
        AddASyncEntry(usParaNr:= SDD_C_ICONT, usRdWr:= 0, dValue:= dValue, pThisObj:= pThis, usEntry:= 1);
        AddASyncEntry(usParaNr:= SDD_C_IPEAK, usRdWr:= 0, dValue:= dValue, pThisObj:= pThis, usEntry:= 1);
        AddASyncEntry(usParaNr:= SDD_C_IPEAKN, usRdWr:= 0, dValue:= dValue, pThisObj:= pThis, usEntry:= 1);
      end_if;

      if AxSetPara[IDX_VEL_PARA] <> 0 then
        pThis$DINT := AxSetPara[IDX_VEL_PARA];
        AddASyncEntry(usParaNr:= SDD_V_KP, usRdWr:= 0, dValue:= dValue, pThisObj:= pThis, usEntry:= 1);
        AddASyncEntry(usParaNr:= SDD_V_TN, usRdWr:= 0, dValue:= dValue, pThisObj:= pThis, usEntry:= 1);
        AddASyncEntry(usParaNr:= SDD_V_T, usRdWr:= 0, dValue:= dValue, pThisObj:= pThis, usEntry:= 1);
        AddASyncEntry(usParaNr:= SDD_V_T2, usRdWr:= 0, dValue:= dValue, pThisObj:= pThis, usEntry:= 1);
        AddASyncEntry(usParaNr:= SDD_V_FILT, usRdWr:= 0, dValue:= dValue, pThisObj:= pThis, usEntry:= 1);
        AddASyncEntry(usParaNr:= SDD_V_NMAX, usRdWr:= 0, dValue:= dValue, pThisObj:= pThis, usEntry:= 1);
        AddASyncEntry(usParaNr:= SDD_V_KPREL, usRdWr:= 0, dValue:= dValue, pThisObj:= pThis, usEntry:= 1);
      end_if;

      if AxSetPara[IDX_POS_PARA] <> 0 then
        pThis$DINT := AxSetPara[IDX_POS_PARA];
        AddASyncEntry(usParaNr:= SDD_P_KV, usRdWr:= 0, dValue:= dValue, pThisObj:= pThis, usEntry:= 1);
        AddASyncEntry(usParaNr:= SDD_P_SFF, usRdWr:= 0, dValue:= dValue, pThisObj:= pThis, usEntry:= 1);
        AddASyncEntry(usParaNr:= SDD_P_PSCALE, usRdWr:= 0, dValue:= dValue, pThisObj:= pThis, usEntry:= 1);
        AddASyncEntry(usParaNr:= SDD_P_SSCALE, usRdWr:= 0, dValue:= dValue, pThisObj:= pThis, usEntry:= 1);
        AddASyncEntry(usParaNr:= SDD_P_TFF, usRdWr:= 0, dValue:= dValue, pThisObj:= pThis, usEntry:= 1);
        AddASyncEntry(usParaNr:= SDD_P_PEMAX, usRdWr:= 0, dValue:= dValue, pThisObj:= pThis, usEntry:= 1);
        AddASyncEntry(usParaNr:= SDD_P_SMODE, usRdWr:= 0, dValue:= dValue, pThisObj:= pThis, usEntry:= 1);
      end_if;

      if AxSetPara[IDX_FD_PARA] <> 0 then
        pThis$DINT := AxSetPara[IDX_FD_PARA];
        AddASyncEntry(usParaNr:= SDD_F_BW, usRdWr:= 0, dValue:= dValue, pThisObj:= pThis, usEntry:= 1);
        AddASyncEntry(usParaNr:= SDD_F_FF, usRdWr:= 0, dValue:= dValue, pThisObj:= pThis, usEntry:= 1);
        AddASyncEntry(usParaNr:= SDD_F_RK, usRdWr:= 0, dValue:= dValue, pThisObj:= pThis, usEntry:= 1);
      end_if;

      if AxSetPara[IDX_APPLI_PARA] <> 0 then
        pThis$DINT := AxSetPara[IDX_APPLI_PARA];
        AddASyncEntry(usParaNr:= SDD_A_JRATIO, usRdWr:= 0, dValue:= dValue, pThisObj:= pThis, usEntry:= 1);
        AddASyncEntry(usParaNr:= SDD_A_VALRT1, usRdWr:= 0, dValue:= dValue, pThisObj:= pThis, usEntry:= 1);
        AddASyncEntry(usParaNr:= SDD_A_VALRT2, usRdWr:= 0, dValue:= dValue, pThisObj:= pThis, usEntry:= 1);
        AddASyncEntry(usParaNr:= SDD_A_VALTT1, usRdWr:= 0, dValue:= dValue, pThisObj:= pThis, usEntry:= 1);
        AddASyncEntry(usParaNr:= SDD_A_VALTT2, usRdWr:= 0, dValue:= dValue, pThisObj:= pThis, usEntry:= 1);
        AddASyncEntry(usParaNr:= SDD_A_CTIME, usRdWr:= 0, dValue:= dValue, pThisObj:= pThis, usEntry:= 1);
        AddASyncEntry(usParaNr:= SDD_A_STIME, usRdWr:= 0, dValue:= dValue, pThisObj:= pThis, usEntry:= 1);
        AddASyncEntry(usParaNr:= SDD_A_STYPE, usRdWr:= 0, dValue:= dValue, pThisObj:= pThis, usEntry:= 1);
        AddASyncEntry(usParaNr:= SDD_A_AVSW, usRdWr:= 0, dValue:= dValue, pThisObj:= pThis, usEntry:= 1);
        AddASyncEntry(usParaNr:= SDD_A_I2TERR, usRdWr:= 0, dValue:= dValue, pThisObj:= pThis, usEntry:= 1);
        AddASyncEntry(usParaNr:= SDD_A_TEMPDE, usRdWr:= 0, dValue:= dValue, pThisObj:= pThis, usEntry:= 1);
        AddASyncEntry(usParaNr:= SDD_A_TEMPMW, usRdWr:= 0, dValue:= dValue, pThisObj:= pThis, usEntry:= 1);
        AddASyncEntry(usParaNr:= SDD_A_STRED, usRdWr:= 0, dValue:= dValue, pThisObj:= pThis, usEntry:= 1);
        AddASyncEntry(usParaNr:= SDD_A_STDT, usRdWr:= 0, dValue:= dValue, pThisObj:= pThis, usEntry:= 1);
        AddASyncEntry(usParaNr:= SDD_A_POS, usRdWr:= 0, dValue:= dValue, pThisObj:= pThis, usEntry:= 1);
        AddASyncEntry(usParaNr:= SDD_A_DNAME1, usRdWr:= 0, dValue:= dValue, pThisObj:= pThis, usEntry:= 1);
        AddASyncEntry(usParaNr:= SDD_A_DNAME2, usRdWr:= 0, dValue:= dValue, pThisObj:= pThis, usEntry:= 1);
        AddASyncEntry(usParaNr:= SDD_A_DNAME3, usRdWr:= 0, dValue:= dValue, pThisObj:= pThis, usEntry:= 1);
        AddASyncEntry(usParaNr:= SDD_A_MODE2, usRdWr:= 0, dValue:= dValue, pThisObj:= pThis, usEntry:= 1);
        AddASyncEntry(usParaNr:= SDD_A_MULTI, usRdWr:= 0, dValue:= dValue, pThisObj:= pThis, usEntry:= 1);
        AddASyncEntry(usParaNr:= SDD_A_CAPREF, usRdWr:= 0, dValue:= dValue, pThisObj:= pThis, usEntry:= 1);
        AddASyncEntry(usParaNr:= SDD_A_EDGE, usRdWr:= 0, dValue:= dValue, pThisObj:= pThis, usEntry:= 1);
        AddASyncEntry(usParaNr:= SDD_A_STTH, usRdWr:= 0, dValue:= dValue, pThisObj:= pThis, usEntry:= 1);
        AddASyncEntry(usParaNr:= SDD_A_INT1, usRdWr:= 0, dValue:= dValue, pThisObj:= pThis, usEntry:= 1);
        AddASyncEntry(usParaNr:= SDD_A_INT2, usRdWr:= 0, dValue:= dValue, pThisObj:= pThis, usEntry:= 1);
        AddASyncEntry(usParaNr:= SDD_A_ICOM, usRdWr:= 0, dValue:= dValue, pThisObj:= pThis, usEntry:= 1);
        AddASyncEntry(usParaNr:= SDD_A_ICOMP, usRdWr:= 0, dValue:= dValue, pThisObj:= pThis, usEntry:= 1);
        AddASyncEntry(usParaNr:= SDD_A_CMIN, usRdWr:= 0, dValue:= dValue, pThisObj:= pThis, usEntry:= 1);
        AddASyncEntry(usParaNr:= SDD_A_BIQCF, usRdWr:= 0, dValue:= dValue, pThisObj:= pThis, usEntry:= 1);
        AddASyncEntry(usParaNr:= SDD_A_BIQFR, usRdWr:= 0, dValue:= dValue, pThisObj:= pThis, usEntry:= 1);
        AddASyncEntry(usParaNr:= SDD_A_BIQCD, usRdWr:= 0, dValue:= dValue, pThisObj:= pThis, usEntry:= 1);
        AddASyncEntry(usParaNr:= SDD_A_BIQDR, usRdWr:= 0, dValue:= dValue, pThisObj:= pThis, usEntry:= 1);
        AddASyncEntry(usParaNr:= SDD_A_CAPFT, usRdWr:= 0, dValue:= dValue, pThisObj:= pThis, usEntry:= 1);
        AddASyncEntry(usParaNr:= SDD_A_ACME, usRdWr:= 0, dValue:= dValue, pThisObj:= pThis, usEntry:= 1);
      end_if;

      if AxSetPara[IDX_ERRORHANDLING] <> 0 then
        pThis$DINT := AxSetPara[IDX_ERRORHANDLING];
        AddASyncEntry(usParaNr:= SDD_I_STATUS, usRdWr:= 0, dValue:= dValue, pThisObj:= pThis, usEntry:= 1);
        AddASyncEntry(usParaNr:= SDD_I_DERROR, usRdWr:= 0, dValue:= dValue, pThisObj:= pThis, usEntry:= 1);
      end_if;

      // get the number of parameters in the drive (only to know if we are at the end of the reading process
      AddASyncEntry(usParaNr:= 0, usRdWr:= 0, dValue:= dValue, pThisObj:= NIL, usEntry:= 2);
      ParaReadCmdAx := 4;
    4 :

      if bdSettings.bReadAxFin = TRUE then
      // wait until the last entry is send the value back

        // now save all parameters in the SRAM / FILE
        if DriveInitType = _SDDRAMEX then
          pSDDData$^void := DriveAxisSet.GetMemPtr();
          DriveAxisSet.SaveRamExData(pData:= pSDDData, udLen:= pSDDData^.udLen, udOffset:= 0);

        elsif DriveInitType = _SDDFILE then
          pSDDData$^void := DriveAxisSet.GetMemPtr();
          DriveAxisSet.SaveRamFileData(pData:= pSDDData, udLen:= pSDDData^.udLen, udOffset:= 0);

        end_if;
        ParaReadCmdAx := 0;

      end_if;
    end_case;
  end_if;

END_FUNCTION

FUNCTION VIRTUAL GLOBAL _DriveAxisBase::SetAbsolutePosition
	VAR_INPUT
		AbsPosition 	: DINT;
	END_VAR
	VAR_OUTPUT
		retcode 	: DINT;
	END_VAR

  retcode := 1;
  if IsOnline() = FALSE then
    retcode := -1;  // no communication available or the initialisation isn't finished
    return;
  end_if;

  //Check if operation is already in progress
  if bdSettings.bSetAbsPos = true then
    retcode := -2;
    return;
  end_if;

  // check if the axis is with an absolute encoder
  if (bdSettings.bNoAbsEnc = FALSE) then
    // if any axis is enabled, the parameter K-FBRW cannot be written
    if DriveMng.IsAnyAxisEnabled() then
      retcode := -4;
      return;
    end_if;

    // set the value of the parameter A-MULTI to 1
    AddASyncEntry(SDD_A_MULTI, 1, 1, this, 0);
    // set the new position to the parameter
    AddASyncEntry(SDD_A_POS, 1, AbsPosition, this, 1);
    // marry the motor with the Drive
    AddASyncEntry(SDD_K_FBRW, 1, 3, this, 1);

    bdSettings.bSetAbsPos := TRUE;
  else
    retcode := -3; // no absolute encoder available
  end_if;

END_FUNCTION

FUNCTION VIRTUAL GLOBAL _DriveAxisBase::SetAbsolutePositionEncoder
	VAR_INPUT
		AbsPosition 	: DINT;
	END_VAR
	VAR_OUTPUT
		retcode 	: DINT;
	END_VAR

  //Init Returncode
  retcode := true;

  //Check if Drive is Online and the Initialization is finished
  if IsOnline() = false then
    retcode := -1;
    return;
  end_if;

  //Check if operation is already in progress
  if bdSettings.bSetAbsPosEncoder = true then
    retcode := -2;
    return;
  end_if;

  //Check if the Axis got an AbsoluteEncoder
  if bdSettings.bNoAbsEnc = false then
    // if axis is enabled, the parameter K-FBRW cannot be written
    if DriveMng.IsAnyAxisEnabled() then
      retcode := -4;
      return;
    end_if;

    //Set A-MULTI to 1
    AddASyncEntry(SDD_A_MULTI, true, 0, this, 0);

    //Set A-POS to InputParamter
    AddASyncEntry(SDD_A_POS, true, AbsPosition, this, 1);

    //Set K-FBRW to 5 => Calculate Offset
    AddASyncEntry(SDD_K_FBRW, true, 5, this, 1);

    //Set K-FBRW to 2 => Save Offset in Feedback
    AddASyncEntry(SDD_K_FBRW, true, 2, this, 1);

    bdSettings.bSetAbsPosEncoder := true;
  else
    retcode := -3;
  end_if;

END_FUNCTION

FUNCTION _DriveAxisBase::SaveDrivePara
  VAR
    TabAddress 	: ^DINT;
    pHlpSDD		: ^void;
    TabLength   : DINT;
  END_VAR

  // get the actual ptr of the memory
  pSDDData$^void := DriveAxisSet.GetMemPtr();

  if pSDDData <> NIL then

    pSDDData^.udLen := sizeof(_SDDMEMHEADER); // initialize the length of the data
    pSDDData^.AxOffset := sizeof(_SDDMEMHEADER); // set the offset
    TabAddress := GetTabAdress(1, bdSettings.bSendMPara, #TabLength);

    if TabAddress = NIL then
      return;
    end_if;

    pSDDData^.AxLength := TabLength$UDINT;

    pHlpSDD := pSDDData + pSDDData^.AxOffset;

    _memcpy(pHlpSDD, (TabAddress)$^void, (TabLength)$UDINT);

    pSDDData^.udLen += pSDDData^.AxLength;

    // calculate the crc of the sdd parameters
    pSDDData^.udCRC32 := CalcCRC32((pSDDData + sizeof(UDINT))$^UDINT, pSDDData^.udLen - sizeof(UDINT));

    case DriveInitType of

    _SDDRAMEX :

      // save the data in the ramex
      DriveAxisSet.SaveRamExData(pSDDData, pSDDData^.udLen, 0);

    _SDDFILE :
      // save the data in the ramfile
      DriveAxisSet.SaveRamFileData(pSDDData, pSDDData^.udLen, 0);

    end_case;
  end_if;

END_FUNCTION

FUNCTION _DriveAxisBase::CalcCRC32
	VAR_INPUT
		pData 	: ^UDINT;
		udLen 	: UDINT;
	END_VAR
	VAR_OUTPUT
		CRC32 	: UDINT;
	END_VAR

	CRC32 := coLinker.CRC32(0, pData$^void, udLen);

END_FUNCTION

FUNCTION VIRTUAL GLOBAL _DriveAxisBase::GetZImpulse
	VAR_OUTPUT
		retcode 	: USINT;
	END_VAR

  retcode:=0;

  if ( ( ActPos and maskZImpulse$DINT ) <> oldRevolutions ) then
    retcode := 1;
    oldRevolutions := (ActPos and maskZImpulse$DINT);
  end_if;

END_FUNCTION

FUNCTION VIRTUAL GLOBAL _DriveAxisBase::ZPulsLatch::Read
	VAR_OUTPUT
		output (EAX) 	: DINT;
	END_VAR

  if bOnlineFinished then

    if ZPulsLatch = 0 then
      output := ZPulsLatch := GetZImpulse();
    else
      output := ZPulsLatch;
      ZPulsLatch := 0;
    end_if;

  else
    ZPulsLatch := 0;
    output := ZPulsLatch;
  end_if;

END_FUNCTION

FUNCTION _DriveAxisBase::SetZPulseMask

  maskZImpulse:=16#FFFFFFFF;
  maskZImpulse:=maskZImpulse SHL (32-ppscale);

  //P-PSCALE  0: 00000000 00000000 00000000 00000000
  //P-PSCALE 10: 11111111 11000000 00000000 00000000
  //P-PSCALE 16: 11111111 11111111 00000000 00000000

END_FUNCTION

FUNCTION VIRTUAL GLOBAL _DriveAxisBase::GetSyncEntry
	VAR_INPUT
		usValue 	: USINT;
		usPData 	: ^DINT;
	END_VAR
	VAR_OUTPUT
		retcode 	: DINT;
	END_VAR

  retcode:=DriveMng.GetSyncEntry(usAxis:=usAxisIndex, usValue:=usValue, usPData:=usPData);

END_FUNCTION

FUNCTION VIRTUAL GLOBAL _DriveAxisBase::AddSyncEntry
	VAR_INPUT
		pThis 	: ^void;
	END_VAR
	VAR_OUTPUT
		retcode 	: BOOL;
	END_VAR

  retcode := FALSE;

  if pThis <> NIL then
    SyncParaObject := pThis$DINT;
    retcode := TRUE;
  end_if;

END_FUNCTION

FUNCTION VIRTUAL GLOBAL _DriveAxisBase::SetSyncEntry
	VAR_INPUT
		usValue 	: USINT;
		usPData 	: DINT;
	END_VAR
	VAR_OUTPUT
		retcode 	: DINT;
	END_VAR

  retcode:=DriveMng.SetSyncEntry(usAxis:=usAxisIndex, usValue:=usValue, usPData:=usPData);

END_FUNCTION

FUNCTION _DriveAxisBase::RefreshIASP
	VAR_INPUT
		Para 	  : DINT;
		Value 	: DINT;
	END_VAR
  VAR
  	UserPara      : CmdStruct;
    UserResult    : Results;
  END_VAR

  // if there is a change in the following values, first we set the pointers to zero, and then we initialize them, allready with the new value

  if AxEnable = 0 then //just do some changes when the axis does not run
    case Para of
      SDD_A_VALTT1:

        _memset(#SyncPara.ActCurrent,0,sizeof(SyncPara.ActCurrent));
        _memset(#SyncPara.ActPos,    0,sizeof(SyncPara.ActPos));
        _memset(#SyncPara.ActSpeed,  0,sizeof(SyncPara.ActSpeed));
        _memset(#SyncPara.Xw,        0,sizeof(SyncPara.Xw));
        _memset(#SyncPara.StateWord, 0,sizeof(SyncPara.StateWord));
        _memset(#SyncPara.DigInputs, 0,sizeof(SyncPara.DigInputs));

        ActValues[0] := to_usint( Value AND 16#000000FF);
        ActValues[1] := to_usint((Value AND 16#0000FF00) SHR 8);

        GetSynchronPara();

      SDD_A_VALTT2:

        _memset(#SyncPara.ActCurrent,0,sizeof(SyncPara.ActCurrent));
        _memset(#SyncPara.ActPos,    0,sizeof(SyncPara.ActPos));
        _memset(#SyncPara.ActSpeed,  0,sizeof(SyncPara.ActSpeed));
        _memset(#SyncPara.Xw,        0,sizeof(SyncPara.Xw));
        _memset(#SyncPara.StateWord, 0,sizeof(SyncPara.StateWord));
        _memset(#SyncPara.DigInputs, 0,sizeof(SyncPara.DigInputs));

        ActValues[2] := to_usint( Value AND 16#000000FF);
        ActValues[3] := to_usint((Value AND 16#0000FF00) SHR 8);
        ActValues[4] := to_usint((Value AND 16#00FF0000) SHR 16);

        if (AxisExtend = 1) & (SyncParaObject<>NIL) then
          UserPara.uiCmd := 10;
          UserPara.aPara[2]:=ActValues[2];
          UserPara.aPara[3]:=ActValues[3];
          UserPara.aPara[4]:=ActValues[4];
          SyncParaObject$^VirtualBase^.pSvrChCmd.NewInst(#UserPara, #UserResult); //initialize also the extend class
        end_if;

        GetSynchronPara();

      SDD_A_VALRT1:

        _memset(#SyncPara.SetCurrent, 0,sizeof(SyncPara.SetCurrent));
        _memset(#SyncPara.SetPos,     0,sizeof(SyncPara.SetPos));
        _memset(#SyncPara.SetSpeed,   0,sizeof(SyncPara.SetSpeed));
        _memset(#SyncPara.SetTorque,  0,sizeof(SyncPara.SetTorque));
        _memset(#SyncPara.ControlWord,0,sizeof(SyncPara.ControlWord));

        SetValues[0] := to_usint( Value AND 16#000000FF);
        SetValues[1] := to_usint((Value AND 16#0000FF00) SHR 8);

        SetSynchronPara();
//        AxTorqueControl.Write(4500); //it does not matter which controlword we have, because the internal function reduced this amount to the top limit
        SetAxTorque(4500);

      SDD_A_VALRT2:

        _memset(#SyncPara.SetCurrent, 0,sizeof(SyncPara.SetCurrent));
        _memset(#SyncPara.SetPos,     0,sizeof(SyncPara.SetPos));
        _memset(#SyncPara.SetSpeed,   0,sizeof(SyncPara.SetSpeed));
        _memset(#SyncPara.SetTorque,  0,sizeof(SyncPara.SetTorque));
        _memset(#SyncPara.ControlWord,0,sizeof(SyncPara.ControlWord));

        SetValues[2] := to_usint( Value AND 16#000000FF);
        SetValues[3] := to_usint((Value AND 16#0000FF00) SHR 8);
        SetValues[4] := to_usint((Value AND 16#00FF0000) SHR 16);

        if (AxisExtend = 1) & (SyncParaObject<>NIL) then
          UserPara.uiCmd := 11;
          UserPara.aPara[2]:=SetValues[2];
          UserPara.aPara[3]:=SetValues[3];
          UserPara.aPara[4]:=SetValues[4];
          SyncParaObject$^VirtualBase^.pSvrChCmd.NewInst(#UserPara, #UserResult); //if there is a extend class connected, we have to initialize it
        end_if;

        SetSynchronPara();
//        AxTorqueControl.Write(4500); //it does not matter which controlword we have, because the internal function reduced this amount to the top limit
        SetAxTorque(4500);

      SDD_P_PSCALE:
        ppscale:=to_usint(Value);
        SetZPulseMask();

    end_case;
  end_if;

END_FUNCTION

FUNCTION VIRTUAL GLOBAL _DriveAxisBase::AxOkay
	VAR_OUTPUT
		retcode 	: DINT;
	END_VAR

  retcode := false;
  if AxisState = 0 then
    retcode := true;
  end_if;

END_FUNCTION

FUNCTION VIRTUAL GLOBAL _DriveAxisBase::Online::Read
	VAR_OUTPUT
		output (EAX) 	: DINT;
	END_VAR

  //--- if DriveMng is online, we have no internal error, and the error-reset after startup is ready, we say Online = 1
//  Online := bOnlineFinished;
  Online := bOnlineState;

  output := Online;

END_FUNCTION

FUNCTION VIRTUAL GLOBAL _DriveAxisBase::ErrorQuitHandling
	VAR_INPUT
		input 	: DINT;
	END_VAR
	VAR_OUTPUT
		result 	: DINT;
	END_VAR

  AxErrorQuit:=input AND 1;

  // check if there is a control word mapped, before accessing the data
  if SyncPara.ControlWord.ptr then
    if (SyncPara.ControlWord.userinfo=0) then
      SyncPara.ControlWord.ptr^$BINT.2:=AxErrorQuit$BOOL; //FAULT RESET
    elsif(SyncPara.ControlWord.userinfo=1) then
      SyncPara.ControlWord.ptr^$BINT.8:=AxErrorQuit$BOOL; //FAULT RESET
    end_if;
  end_if;

  if AxErrorQuit = 1 then
    FirstErrorReset := 4;
    ErrorQuitTime:=ops.tAbsolute;
  end_if;

  Controlword.ResetFault := AxErrorQuit$BOOL;

  result := AxErrorQuit;

END_FUNCTION

FUNCTION VIRTUAL _DriveAxisBase::GetAxError
	VAR_OUTPUT
		AxError 	: DINT;
	END_VAR
  VAR
  	sBuffer      : BDINT; //StateWord Buffer
  END_VAR

  if SyncPara.StateWord.ptr<>NIL  then
    sBuffer := SyncPara.StateWord.ptr^$BDINT;
    AxError:=sBuffer.4; //the error is at both control words on the same place
  else
    AxError:=0;
  end_if;

END_FUNCTION

FUNCTION _DriveAxisBase::SetAxTorque
	VAR_INPUT
		NewTorque 	: UDINT;
	END_VAR
  VAR
    cBuffer       : BDINT; //ControlWord Buffer
  END_VAR

  // if we have a 16-Bit Controlword
  if SyncPara.SetTorque.userinfo = 0 then

    if NewTorque < 0 then
      NewTorque := 0;
    end_if;

    if NewTorque > DRIVEAXIS_TORQUE_LIMITATION_VALUE then
      NewTorque := DRIVEAXIS_TORQUE_LIMITATION_VALUE;
    end_if;

    AxTorqueControl := NewTorque;

    //Check if pointer is valid
    if SyncPara.ControlWord.ptr then
      cBuffer:=SyncPara.ControlWord.ptr^$BDINT;
      SyncPara.SetTorque.ptr^$INT:= to_int(TorqueCalculation(cBuffer,NewTorque));
    end_if;

  elsif SyncPara.SetTorque.userinfo=1 then //that is for the 32-Bit Controlword

    if NewTorque < 0 then
      NewTorque := 0;
    end_if;

    if NewTorque > 4500 then
      NewTorque := 4500;
    end_if;

    AxTorqueControl := NewTorque;

    if SyncPara.SetTorque.ptr then
      SyncPara.SetTorque.ptr^$INT:=to_int(NewTorque);
    end_if;

  end_if;

END_FUNCTION

FUNCTION _DriveAxisBase::IsOnlineFinished
	VAR_OUTPUT
		bOnline 	: BOOL;
	END_VAR

  if (IsOnline() = TRUE) & (CmdState <> ERROR) & ((FirstErrorReset = 0) | (FirstErrorReset >= 4)) then
    bOnline := 1;
  else
    bOnline := 0;
  end_if;

END_FUNCTION

FUNCTION VIRTUAL GLOBAL _DriveAxisBase::AddASyncEntryDS402
	VAR_INPUT
		uiParaID 	  : UINT;
		usParaSubID : USINT;
		usRdWr 	    : USINT;
		pValue 	    : ^USINT;
		bsDataInfo 	: BSINT;
		pThisObj 	  : ^void;
		usEntry 	  : USINT;
	END_VAR
	VAR_OUTPUT
		retcode 	  : DINT;
	END_VAR

  retcode := DriveMng.AddASyncEntryDS402(AxisNo     := usAxisIndex
                                      , uiParaID    := uiParaID
                                      , usParaSubID := usParaSubID
                                      , usRdWr      := usRdWr
                                      , pValue      := pValue
                                      , bsDataInfo  := bsDataInfo
                                      , pThisObj    := pThisObj
                                      , usEntry     := usEntry
                                      );

END_FUNCTION

FUNCTION VIRTUAL GLOBAL _DriveAxisBase::Input1::Read
	VAR_OUTPUT
		output (EAX) 	: DINT;
	END_VAR

  if (SyncPara.DigInputs.ptr <> NIL) & bOnlineFinished then
    if SyncPara.DigInputs.size >= 1 then
      Input1:=SyncPara.DigInputs.ptr^$BSINT.1;
    else
      Input1:=0;
    end_if;
  else
    Input1:=0;
  end_if;

	output := Input1;

END_FUNCTION

FUNCTION VIRTUAL GLOBAL _DriveAxisBase::Input2::Read
	VAR_OUTPUT
		output (EAX) 	: DINT;
	END_VAR

  if (SyncPara.DigInputs.ptr <> NIL) & bOnlineFinished then
    if SyncPara.DigInputs.size >= 2 then
      Input2:=SyncPara.DigInputs.ptr^$BSINT.2;
    else
      Input2:=0;
    end_if;
  else
    Input2:=0;
  end_if;

	output := Input2;

END_FUNCTION

FUNCTION VIRTUAL GLOBAL _DriveAxisBase::Input3::Read
	VAR_OUTPUT
		output (EAX) 	: DINT;
	END_VAR

  if (SyncPara.DigInputs.ptr <> NIL) & bOnlineFinished then
    if SyncPara.DigInputs.size >= 3 then
      Input3:=SyncPara.DigInputs.ptr^$BSINT.3;
    else
      Input3:=0;
    end_if;
  else
    Input3:=0;
  end_if;

	output := Input3;

END_FUNCTION

FUNCTION VIRTUAL GLOBAL _DriveAxisBase::Input4::Read
	VAR_OUTPUT
		output (EAX) 	: DINT;
	END_VAR

  if (SyncPara.DigInputs.ptr <> NIL) & bOnlineFinished then
    if SyncPara.DigInputs.size >= 4 then
      Input4:=SyncPara.DigInputs.ptr^$BSINT.4;
    else
      Input4:=0;
    end_if;
  else
    Input4:=0;
  end_if;

	output := Input4;

END_FUNCTION

FUNCTION VIRTUAL GLOBAL _DriveAxisBase::Input5::Read
	VAR_OUTPUT
		output (EAX) 	: DINT;
	END_VAR

  if (SyncPara.DigInputs.ptr <> NIL) & bOnlineFinished then
    if SyncPara.DigInputs.size >= 5 then
      Input5:=SyncPara.DigInputs.ptr^$BSINT.5;
    else
      Input5:=0;
    end_if;
  else
    Input5:=0;
  end_if;

	output := Input5;

END_FUNCTION

FUNCTION VIRTUAL GLOBAL _DriveAxisBase::Input6::Read
	VAR_OUTPUT
		output (EAX) 	: DINT;
	END_VAR

  if (SyncPara.DigInputs.ptr <> NIL) & bOnlineFinished then
    if SyncPara.DigInputs.size >= 6 then
      Input6:=SyncPara.DigInputs.ptr^$BSINT.6;
    else
      Input6:=0;
    end_if;
  else
    Input6:=0;
  end_if;

	output := Input6;

END_FUNCTION

FUNCTION VIRTUAL GLOBAL _DriveAxisBase::Input7::Read
	VAR_OUTPUT
		output (EAX) 	: DINT;
	END_VAR

  if (SyncPara.DigInputs.ptr <> NIL) & bOnlineFinished then
    if SyncPara.DigInputs.size >= 7 then
      Input7:=SyncPara.DigInputs.ptr^$BSINT.7;
    else
      Input7:=0;
    end_if;
  else
    Input7:=0;
  end_if;

	output := Input7;

END_FUNCTION

FUNCTION VIRTUAL GLOBAL _DriveAxisBase::Input8::Read
	VAR_OUTPUT
		output (EAX) 	: DINT;
	END_VAR

  if (SyncPara.DigInputs.ptr <> NIL) & bOnlineFinished then
    if SyncPara.DigInputs.size >= 8 then
      Input8:=SyncPara.DigInputs.ptr^$BSINT.8;
    else
      Input8:=0;
    end_if;
  else
    Input8:=0;
  end_if;

	output := Input8;

END_FUNCTION

FUNCTION VIRTUAL GLOBAL _DriveAxisBase::Output1::Write
	VAR_INPUT
		input (EAX) 	: DINT;
	END_VAR
	VAR_OUTPUT
		result (EAX) 	: DINT;
	END_VAR

  if (SyncPara.ControlWord.ptr <> NIL) & bOnlineFinished then

    if (SyncPara.ControlWord.userinfo=0) then
      Output1 := input AND 1;
      SyncPara.ControlWord.ptr^$BINT.5:=Output1$BOOL; //ManufactureSpec4;  //Output1
      Controlword.ManufactureSpec4 := Output1$BOOL;
    elsif(SyncPara.ControlWord.userinfo=1) then
      //not available in 32bit controlword
      Output1 := 0;
    end_if;

  end_if;

	result := Output1;

END_FUNCTION

FUNCTION VIRTUAL GLOBAL _DriveAxisBase::Output2::Write
	VAR_INPUT
		input (EAX) 	: DINT;
	END_VAR
	VAR_OUTPUT
		result (EAX) 	: DINT;
	END_VAR

  if (SyncPara.ControlWord.ptr <> NIL) & bOnlineFinished then

    if (SyncPara.ControlWord.userinfo=0) then
      Output2 := input AND 1;
      SyncPara.ControlWord.ptr^$BINT.6:=Output2$BOOL; //ManufactureSpec5;  //Output2
      Controlword.ManufactureSpec5 := Output2$BOOL;
    elsif(SyncPara.ControlWord.userinfo=1) then
      //not available in 32bit controlword
      Output2 := 0;
    end_if;

  end_if;

	result := Output2;

END_FUNCTION

#pragma warning(disable: 73);
FUNCTION VIRTUAL _DriveAxisBase::LogError
	VAR_INPUT
		pMsg 	: ^CHAR;
	END_VAR

#ifdef HWC_LogError
  HWC_LogError(this, pMsg);
#endif

END_FUNCTION

FUNCTION VIRTUAL _DriveAxisBase::LogValue
	VAR_INPUT
		pString 	: ^CHAR;
		udValue 	: UDINT;
		udValue2 	: UDINT;(* := 16#FFFFFFFF *)
		udValue3 	: UDINT;(* := 16#FFFFFFFF *)
	END_VAR

#ifdef HWC_LogValue3
  HWC_LogValue3(this, pString, udValue, udValue2, udValue3);
#endif

END_FUNCTION
#pragma warning(default: 73);

FUNCTION GLOBAL _DriveAxisBase::SetDiagMode
	VAR_INPUT
		bStartDiagMode 	: BOOL;
		pThisObj 	: ^void;
	END_VAR
	VAR_OUTPUT
		dRetCode 	: DINT;
	END_VAR

  // initialize return code with ok
  dRetCode := 1;
  if pThisObj <> NIL then
    if bStartDiagMode = TRUE then
      if AxisState.DiagModeActive = FALSE then
        if bOnlineFinished = TRUE then
          AxisState.DiagModeActive := TRUE;
          pDiagThis       := pThisObj;
          bOnlineFinished := FALSE;
        else
          //axis is not online or init is not finished
          dRetCode := -1;
        end_if;
      else
        if pThisObj <> pDiagThis then
          //diag mode is already set by other instance
          dRetCode := -2;
        end_if;
      end_if;

    else
      if pThisObj = pDiagThis then
        //diag mode is deactivated - reset values
        AxisState.DiagModeActive := FALSE;
        pDiagThis := NIL;
        //set act state
        bOnlineFinished := IsOnlineFinished();
      else
        //class was locked by other object
        dRetCode := -3;
      end_if;
    end_if;
  else
    //this pointer is not valid
    dRetCode := -4;
  end_if;

END_FUNCTION

FUNCTION GLOBAL _DriveAxisBase::GetDriveType
	VAR_OUTPUT
		DriveType 	: _DRIVETYPE;
	END_VAR

  DriveType := DriveMng.DriveType;

END_FUNCTION

FUNCTION _DriveAxisBase::Write_SetSpeed
	VAR_INPUT
		valueIn 	: DINT;
	END_VAR
	VAR_OUTPUT
		valueOut 	: DINT;
	END_VAR

  // writes the value to the PDO data.
  // online is not checked on purpose. It is needed to initialize the PDO data for a reconnect.
  // The value may be truncated to 16bit in the PDO, but is not for the return value.

  valueOut := 0;// zero in case we have no access
	if (SyncPara.SetSpeed.ptr <> NIL) then

    if (SyncPara.SetSpeed.size=4) then
      SyncPara.SetSpeed.ptr^ := valueIn;
      valueOut := valueIn;

    elsif (SyncPara.SetSpeed.size=2) then
      if SyncPara.SetSpeed.userinfo = 0 then
        if valueIn > DRIVEAXIS_SPEED_SFFLIMITATION_USERINFO_0 then
          valueIn := DRIVEAXIS_SPEED_SFFLIMITATION_USERINFO_0;
          AxisState.SFFLimitationActive := TRUE;
        elsif valueIn < -DRIVEAXIS_SPEED_SFFLIMITATION_USERINFO_0-1 then
          valueIn := -DRIVEAXIS_SPEED_SFFLIMITATION_USERINFO_0-1;
          AxisState.SFFLimitationActive := TRUE;
        else
          AxisState.SFFLimitationActive := FALSE;
        end_if;
        SyncPara.SetSpeed.ptr^$INT := to_int(valueIn);
        valueOut := valueIn;
      elsif SyncPara.SetSpeed.userinfo = 1 then
        if valueIn > DRIVEAXIS_SPEED_SFFLIMITATION_USERINFO_1 then
          valueIn := DRIVEAXIS_SPEED_SFFLIMITATION_USERINFO_1;
          AxisState.SFFLimitationActive := TRUE;
        elsif valueIn < -DRIVEAXIS_SPEED_SFFLIMITATION_USERINFO_1 then
          valueIn := -DRIVEAXIS_SPEED_SFFLIMITATION_USERINFO_1;
          AxisState.SFFLimitationActive := TRUE;
        else
          AxisState.SFFLimitationActive := FALSE;
        end_if;
        SyncPara.SetSpeed.ptr^$INT := to_int(valueIn);
        valueOut := valueIn;
      end_if;
    end_if;
  end_if;

END_FUNCTION

FUNCTION _DriveAxisBase::Write_Enable
	VAR_INPUT
		valueIn 	: DINT;
	END_VAR
	VAR_OUTPUT
		valueOut 	: DINT;
	END_VAR

  // writes the value to the PDO data.
  // online is not checked on purpose. It is needed to initialize the PDO data for a reconnect.

  valueOut := 0;// zero in case we have no access
  if (SyncPara.ControlWord.ptr <> NIL) then
    if (SyncPara.ControlWord.userinfo=0) then
      SyncPara.ControlWord.ptr^$BINT.1:=valueIn$BOOL; //DRIVE ENABLE
    elsif(SyncPara.ControlWord.userinfo=1) then
      SyncPara.ControlWord.ptr^$BINT.4:=valueIn$BOOL; //DRIVE ENABLE
    end_if;

    Controlword.EnableOperation := valueIn$BOOL;
    valueOut := to_dint(valueIn$BOOL);
  end_if;

END_FUNCTION
